Omron CX-Programmer project NewProject (CX-Programmer 9.61)

# PLC NewPLC1: CJ1M CPU21

## Global symbols (name address type ; comment)
Humidity_1 Humidity
K K1
Temperature Temperature
Temperature_0 Temperature
Temperature_1 Temperature
Temperature_2 Temperature
Temperature_3 Temperature

## Program НоваяЗадача1 (cyclic task 0)

### Section Сегмент1

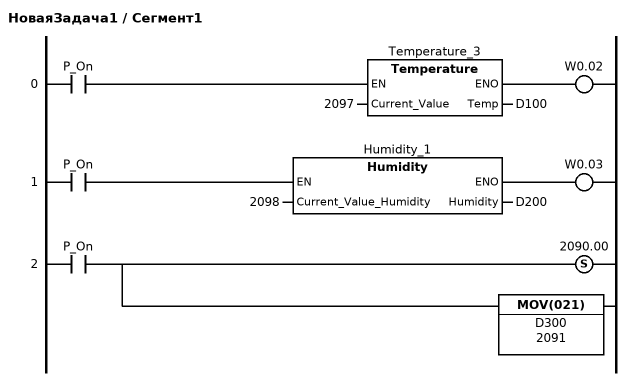
; rung 0
LD P_On
CALL Temperature_3 : Temperature (Current_Value := 2097, Temp => D100)
OUT W0.02
; rung 1
LD P_On
CALL Humidity_1 : Humidity (Current_Value_Humidity := 2098, Humidity => D200)
OUT W0.03
; rung 2
LD P_On
SET 2090.00
MOV(021) D300 2091

### Section END
; rung 0
END(001)

## Function block Humidity
VAR_INPUT
  Current_Value_Humidity : INT;
END_VAR
VAR_OUTPUT
  Humidity : REAL;
END_VAR
VAR
  IHumid : REAL;
  Real_Value_Humidity : REAL;
END_VAR
Real_Value_Humidity:= INT_TO_REAL(Current_Value_Humidity);
IHumid:= (Real_Value_Humidity/250.0)+4.0;
Humidity:= (IHumid-4.0)/16.0*95.0;

## Function block Temperature
VAR_INPUT
  Current_Value : INT;
END_VAR
VAR_OUTPUT
  Temp : REAL;
END_VAR
VAR
  Itemp : REAL;
  Real_Current_Value : REAL;
END_VAR
Real_Current_Value:= INT_TO_REAL(Current_Value);
Itemp:= 4.0 + (Real_Current_Value / 4000.0) * 16.0;
Temp:= ((Itemp-4.0)/16.0)*90.0-20.0;